// TIA Portal V20 program export: 1 tag tables, 0 data types, 1 data blocks, 2 code blocks (in call order from the OBs), 1 instance data blocks

VAR_GLOBAL   // PLC tag table "Cinta_Signals"
   DI_ES01_Ok AT %M0.0 : Bool;
   DI_M01_Start AT %M0.1 : Bool;
   DI_M01_Stop AT %M0.2 : Bool;
   DI_M01_Reset AT %M0.3 : Bool;
   DI_M01_Feedback AT %M0.4 : Bool;
   DO_M01_Run AT %M1.0 : Bool;
   M_M01_Running AT %M1.1 : Bool;
   M_M01_Interlock AT %M1.2 : Bool;
   M_M01_Fault AT %M1.3 : Bool;
   M_M01_FaultCode AT %MW4 : Int;
END_VAR

// Al generar este bloque, TIA crea el DB de instancia "iDB_M01" del FB_Motor.
//==============================================================================
DATA_BLOCK "iDB_M01"
{ S7_Optimized_Access := 'TRUE' }
VERSION : 0.1
   "FB_Motor"
END_DATA_BLOCK

ORGANIZATION_BLOCK "Main"
{ S7_Optimized_Access := 'TRUE' }
VERSION : 0.1
AUTHOR : JMellid
FAMILY : Drives
//==============================================================================
// OB ciclico de la cinta DEMO-Cinta01.
//
// El OB ciclico se llama "Main" porque ese es el nombre que le pone TIA al
// OB1 del sistema: generar desde una fuente un OB llamado "OB_Main" falla con
// 'Type conflict: Object "OB_Main" cannot be overwritten'. El estandar
// OB_<Funcion> de 20-standards/naming.md aplica a los OB de arranque y de
// error, no al OB1 del sistema, cuyo nombre es de TIA.
//
// Una cinta con un solo motor (M01) y seta de emergencia.
//
// El enclavamiento NO se calcula dentro del FB: se ve aqui, en el punto de
// llamada, que es donde lo mira el mantenedor de la maquina. Ver R08.
//
// La seta de emergencia (DI_ES01_Ok, contacto normalmente cerrado: TRUE cuando
// NO esta pulsada) hace las dos cosas que tiene que hacer, y las dos son
// obligatorias:
//   1. Prohíbe arrancar: el Interlock del FB exige DI_ES01_Ok.
//   2. Ordena parar:     CmdStop incluye NOT DI_ES01_Ok, de modo que con la
//                        seta pulsada el motor para aunque nadie pulse el
//                        boton de paro.
// Si solo se hiciera la primera, el motor seguiria girando con la seta
// pulsada. Eso no es una seta de emergencia: es un pulsador de arranque.
//
// "DI_M01_Start" y "DI_M01_Stop" los escribe el HMI (botones de la pantalla
// Main) y tambien pueden venir de un pulsador de campo. "DI_M01_Feedback"
// llega del contacto auxiliar del contactor.
//
// Al generar este bloque, TIA crea el DB de instancia "iDB_M01" del FB_Motor.
//==============================================================================
BEGIN
   "iDB_M01"(CmdStart     := "DI_M01_Start",
             CmdStop      := "DI_M01_Stop" OR NOT "DI_ES01_Ok",
             CmdReset     := "DI_M01_Reset",
             Interlock    := "DI_ES01_Ok",
             Feedback     := "DI_M01_Feedback",
             FeedbackUsed := TRUE,
             StartTimeout := T#3S,
             StopTimeout  := T#3S,
             Run          => "DO_M01_Run",
             Running      => "M_M01_Running",
             Ready        => "M_M01_Interlock",
             Fault        => "M_M01_Fault",
             FaultCode    => "M_M01_FaultCode");
END_ORGANIZATION_BLOCK

ORGANIZATION_BLOCK "Main"   // OB1, SCL, ProgramCycle
{ S7_Optimized_Access := 'TRUE' }
AUTHOR : JMellid
FAMILY : Drives
// ==============================================================================
//  OB ciclico de la cinta DEMO-Cinta01.
// 
//  El OB ciclico se llama "Main" porque ese es el nombre que le pone TIA al
//  OB1 del sistema: generar desde una fuente un OB llamado "OB_Main" falla con
//  'Type conflict: Object "OB_Main" cannot be overwritten'. El estandar
//  OB_<Funcion> de 20-standards/naming.md aplica a los OB de arranque y de
//  error, no al OB1 del sistema, cuyo nombre es de TIA.
// 
//  Una cinta con un solo motor (M01) y seta de emergencia.
// 
//  El enclavamiento NO se calcula dentro del FB: se ve aqui, en el punto de
//  llamada, que es donde lo mira el mantenedor de la maquina. Ver R08.
// 
//  La seta de emergencia (DI_ES01_Ok, contacto normalmente cerrado: TRUE cuando
//  NO esta pulsada) hace las dos cosas que tiene que hacer, y las dos son
//  obligatorias:
//    1. ProhÃ­be arrancar: el Interlock del FB exige DI_ES01_Ok.
//    2. Ordena parar:     CmdStop incluye NOT DI_ES01_Ok, de modo que con la
//                         seta pulsada el motor para aunque nadie pulse el
//                         boton de paro.
//  Si solo se hiciera la primera, el motor seguiria girando con la seta
//  pulsada. Eso no es una seta de emergencia: es un pulsador de arranque.
// 
//  "DI_M01_Start" y "DI_M01_Stop" los escribe el HMI (botones de la pantalla
//  Main) y tambien pueden venir de un pulsador de campo. "DI_M01_Feedback"
//  llega del contacto auxiliar del contactor.
// 
//  Al generar este bloque, TIA crea el DB de instancia "iDB_M01" del FB_Motor.
// ==============================================================================
// stored: SetENOAutomatically false
   VAR_INPUT
      Initial_Call : Bool;   // Initial call of this OB
      Remanence : Bool;   // =True, if remanent data are available
   END_VAR
BEGIN

   "iDB_M01"(CmdStart := "DI_M01_Start",
             CmdStop := "DI_M01_Stop" OR NOT "DI_ES01_Ok",
             CmdReset := "DI_M01_Reset",
             Interlock := "DI_ES01_Ok",
             Feedback := "DI_M01_Feedback",
             FeedbackUsed := TRUE,
             StartTimeout := T#3S,
             StopTimeout := T#3S,
             Run => "DO_M01_Run",
             Running => "M_M01_Running",
             Ready => "M_M01_Interlock",
             Fault => "M_M01_Fault",
             FaultCode => "M_M01_FaultCode");
END_ORGANIZATION_BLOCK

FUNCTION_BLOCK "FB_Motor"   // FB1, SCL
{ S7_Optimized_Access := 'TRUE' }
AUTHOR : JMellid
FAMILY : Drives
// ==============================================================================
//  Mando de un motor de marcha/paro con confirmacion y deteccion de fallo.
// 
//  Arranca con CmdStart si Interlock lo permite. Si no llega Feedback antes de
//  StartTimeout, levanta Fault y corta la salida. Si la confirmacion se pierde
//  estando en marcha, tambien. El fallo es enclavado: solo lo borra CmdReset.
// 
//  El enclavamiento NO se calcula aqui: entra por Interlock, para que la cadena
//  de condiciones se vea en LAD en el punto de llamada, que es donde la mira el
//  mantenedor. Ver 10-kb/20-recetas/R08-bloque-motor.md
// ==============================================================================
// stored: MemoryReserve 100, SetENOAutomatically false
   VAR_INPUT
      CmdStart : Bool;   // Orden de marcha (pulso o mantenida)
      CmdStop : Bool;   // Orden de paro. Manda sobre CmdStart
      CmdReset : Bool;   // Rearme del fallo enclavado
      Interlock : Bool := TRUE;   // TRUE = permitido arrancar
      Feedback : Bool;   // Confirmacion de marcha desde campo
      FeedbackUsed : Bool := TRUE;   // FALSE si el motor no tiene retorno
      StartTimeout : Time := T#3S;   // Espera maxima de confirmacion
      StopTimeout : Time := T#3S;   // Espera maxima hasta que cae Feedback
   END_VAR
   VAR_OUTPUT
      Run : Bool;   // Salida al contactor
      Running : Bool;   // Marcha confirmada
      Ready : Bool;   // Disponible para arrancar
      Fault : Bool;   // Fallo enclavado
      FaultCode : Int;   // 0 = sin fallo, ver constantes
   END_VAR
   VAR
      statRunLatch : Bool;   // Memoria de la orden de marcha
      statWasConfirmed : Bool;   // Hubo confirmacion en este arranque
      statFault : Bool;   // Estado interno del fallo
      statFaultCode : Int;   // Codigo interno del fallo
      tonStart { S7_SetPoint := 'True'} : TON_TIME;   // Vigila la aparicion de Feedback
      tonStop { S7_SetPoint := 'True'} : TON_TIME;   // Vigila la desaparicion de Feedback
   END_VAR
   VAR CONSTANT
      FAULT_NONE : Int := 0;
      FAULT_NO_FEEDBACK : Int := 101;   // No confirmo la marcha a tiempo
      FAULT_FEEDBACK_LOST : Int := 102;   // Confirmo y despues se perdio
      FAULT_NO_STOP : Int := 103;   // Sigue confirmando tras el paro
   END_VAR
BEGIN


   REGION 1 - Rearme del fallo
       // Va primero: un rearme debe surtir efecto en el mismo ciclo.
       IF #CmdReset THEN
           #statFault := FALSE;
           #statFaultCode := #FAULT_NONE;
           #statWasConfirmed := FALSE;
       END_IF;
   END_REGION

   REGION 2 - Memoria de marcha
       // El paro, el fallo y el enclavamiento mandan SIEMPRE sobre la orden de
       // marcha. Esta rama va primero para que se falle por el lado seguro.
       IF #CmdStop OR #statFault OR NOT #Interlock THEN
           #statRunLatch := FALSE;
       ELSIF #CmdStart THEN
           #statRunLatch := TRUE;
       END_IF;
   END_REGION

   REGION 3 - Vigilancia de la confirmacion
       // tonStart cubre los dos casos: nunca confirmo, y confirmo y se perdio.
       // La diferencia la da statWasConfirmed, para dar un codigo distinto.
       #tonStart(IN := #statRunLatch AND #FeedbackUsed AND NOT #Feedback,
                 PT := #StartTimeout);

       #tonStop(IN := NOT #statRunLatch AND #FeedbackUsed AND #Feedback,
                PT := #StopTimeout);

       IF #statRunLatch AND #Feedback THEN
           #statWasConfirmed := TRUE;
       END_IF;

       IF NOT #statFault THEN
           IF #tonStart.Q THEN
               #statFault := TRUE;
               IF #statWasConfirmed THEN
                   #statFaultCode := #FAULT_FEEDBACK_LOST;
               ELSE
                   #statFaultCode := #FAULT_NO_FEEDBACK;
               END_IF;
           ELSIF #tonStop.Q THEN
               #statFault := TRUE;
               #statFaultCode := #FAULT_NO_STOP;
           END_IF;
       END_IF;

       IF NOT #statRunLatch THEN
           #statWasConfirmed := FALSE;
       END_IF;
   END_REGION

   REGION 4 - Salidas
       // Cada salida se escribe en UN solo sitio, al final del bloque.
       // El estado vive en variables stat; las salidas solo lo publican.
       // Si se leyera #Fault en la logica, el compilador avisa de que puede no
       // estar inicializado: las salidas se escriben, no se usan como memoria.
       #Run := #statRunLatch AND NOT #statFault;
       #Running := #Run AND (#Feedback OR NOT #FeedbackUsed);
       #Ready := #Interlock AND NOT #statFault AND NOT #statRunLatch;
       #Fault := #statFault;
       #FaultCode := #statFaultCode;
   END_REGION
END_FUNCTION_BLOCK

DATA_BLOCK "iDB_M01"   // DB1
AUTHOR : JMellid
FAMILY : Drives
// Al generar este bloque, TIA crea el DB de instancia "iDB_M01" del FB_Motor.
// ==============================================================================
// stored: InstanceOfName FB_Motor, InstanceOfType FB
"FB_Motor"
BEGIN
END_DATA_BLOCK
